(* PLC project TBEN_L5_PLC11.project, CODESYS CODESYS V3.5 SP21 Patch 1 *)
(* stored: creationDateTime 2026-11-07T15:35:24.8913158, modificationDateTime 2026-11-07T15:09:07.4034196 *)

(* global variable list GVL_IolSys *)
{attribute 'qualified_only'}
// Instance master + transport IO-Link (gọi trong PRG_IOLink / MainTask)
VAR_GLOBAL
    xSimMode  : BOOL := TRUE;              // TRUE = dùng mock (Simulation). Đặt FALSE sau khi có PROFINET thật.
    fbMockAL1 : FB_MockRecordAccess;       // giả lập AL1100 + O5D150
    fbPnAL1   : FB_PnRecordAccess;         // transport PROFINET thật (hiện là khung)
    fbAL1     : FB_IolMaster;              // master AL1100: khoá + hàng đợi IOL_CALL
END_VAR
